(* Logix 5000 project; controller WWTP_CLX vendor 1 type 14 code 54 rev 17.2; software revision 17.00; part 11 of 13 *)

ADD_ON_INSTRUCTION U_FlowTot   (* revision 1.0 *)
// Provides Totalization for Daily & Yearly Flow.
VAR_IN_OUT
   Inp_AIn : P_AIn; {required}   // Flow Analog Input AOI
   Inp_WallClock : U_WallClock; {required}   // PLC Wall Clock
END_VAR
VAR_INPUT
   Inp_ProgStartReq : BOOL := 1;   // Prog Start Request. If needed map to turn on totalizer, (ex. pump running) else Defaults to 1 (always start)
END_VAR
VAR_OUTPUT
   Val_FlowRate : REAL; {visible}   // Current Flow Rate
   Val_DailyTot : REAL; {visible}   // Todays Total Flow
   Val_YestTot : REAL; {visible}   // Yesterday Total Flow
   Val_YearlyTot : REAL; {visible}   // This Year Total Flow
   Val_LastYearTot : REAL; {visible}   // Last Year Total Flow
END_VAR
VAR
   YearlyTotalizer : TOTALIZER := (TimeBase := 3, Gain := 1.0, ProgProgReq := 1, ProgStartReq := 1, OperStartReq := 1, RTSTime := 1, ProgOper := 1, RunStop := 1, TargetFlag := 1, TargetDev1Flag := 1, TargetDev2Flag := 1, DeltaT := 0.010000001);
   DailyTotalizer : TOTALIZER := (TimeBase := 3, Gain := 100000.0, ProgStartReq := 1, OperStartReq := 1, RTSTime := 1, ProgOper := 1, RunStop := 1, TargetFlag := 1, TargetDev1Flag := 1, TargetDev2Flag := 1, DeltaT := 0.010000001);
   FlowRateLowLimit_SSUM : SELECTED_SUMMER := (Gain1 := 1.0, Gain2 := 1.0, Gain3 := 1.0, Gain4 := 1.0, Gain5 := 1.0, Gain6 := 1.0, Gain7 := 1.0, Gain8 := 1.0);
   LowCutoff_BNOT : FBD_BOOLEAN_NOT := (In := 1);
   __l000041A5 : DINT;
   __l000035B4 : REAL;
   __l00000EE7 : BOOL;
   __l00002582 : DINT;
END_VAR

ROUTINE Logic   (* function block diagram *)
   SHEET 1   // Main
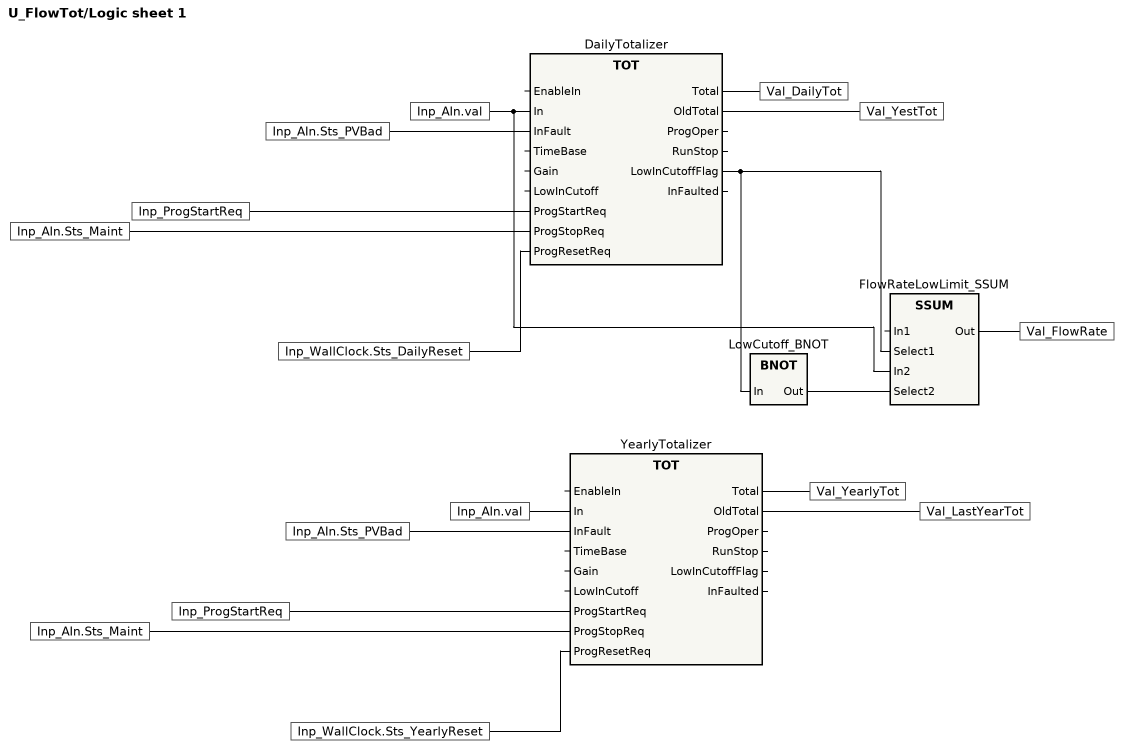
   DailyTotalizer : TOT(In := Inp_AIn.val, InFault := Inp_AIn.Sts_PVBad, ProgStartReq := Inp_ProgStartReq, ProgStopReq := Inp_AIn.Sts_Maint, ProgResetReq := Inp_WallClock.Sts_DailyReset);   // unwired pins: EnableIn TimeBase Gain LowInCutoff ProgOper RunStop InFaulted
   YearlyTotalizer : TOT(In := Inp_AIn.val, InFault := Inp_AIn.Sts_PVBad, ProgStartReq := Inp_ProgStartReq, ProgStopReq := Inp_AIn.Sts_Maint, ProgResetReq := Inp_WallClock.Sts_YearlyReset);   // unwired pins: EnableIn TimeBase Gain LowInCutoff ProgOper RunStop LowInCutoffFlag InFaulted
   LowCutoff_BNOT : BNOT(In := DailyTotalizer.LowInCutoffFlag);
   Val_DailyTot := DailyTotalizer.Total;
   Val_YearlyTot := YearlyTotalizer.Total;
   Val_YestTot := DailyTotalizer.OldTotal;
   FlowRateLowLimit_SSUM : SSUM(Select1 := DailyTotalizer.LowInCutoffFlag, In2 := Inp_AIn.val, Select2 := LowCutoff_BNOT.Out);   // unwired pins: In1
   Val_LastYearTot := YearlyTotalizer.OldTotal;
   Val_FlowRate := FlowRateLowLimit_SSUM.Out;
END_ROUTINE
END_ADD_ON_INSTRUCTION

ADD_ON_INSTRUCTION U_Heartbeat   (* revision 1.0 *)
// Heartbeat Between two PLCs
VAR_INPUT
   CFG_DelayTimerSec : DINT := 30; {visible}   // Delay Timer in Seconds
END_VAR
VAR_OUTPUT
   Heartbeat : BOOL; {visible}   // Heartbeat from Remote PLC
END_VAR
VAR
   DelayTimerOn : TIMER;
   DelayTimerOff : TIMER;
END_VAR

ROUTINE Logic   (* ladder *)
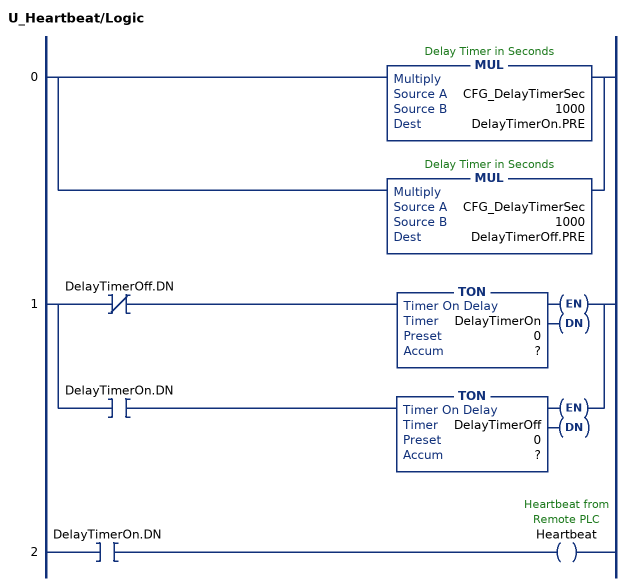
   0: [MUL(CFG_DelayTimerSec,1000,DelayTimerOn.PRE) ,MUL(CFG_DelayTimerSec,1000,DelayTimerOff.PRE) ];
   1: [XIO(DelayTimerOff.DN) TON(DelayTimerOn,?,?) ,XIC(DelayTimerOn.DN) TON(DelayTimerOff,?,?) ];
   2: XIC(DelayTimerOn.DN)OTE(Heartbeat);
END_ROUTINE
END_ADD_ON_INSTRUCTION

ADD_ON_INSTRUCTION U_Module   (* revision 1.0 *)
VAR_INPUT
   EntryStatus : INT; {visible}   // Module Entry Status
   CommLossTimerPresetSec : REAL; {visible}   // Communication Loss Timer Preset (Sec)
END_VAR
VAR_OUTPUT
   CommLoss : BOOL; {visible}   // Communication Loss Alarm
END_VAR
VAR
   ConnectionStatus : DINT;
   CommLossTimer : TIMER := (PRE := 5);
END_VAR

ROUTINE Logic   (* ladder *)
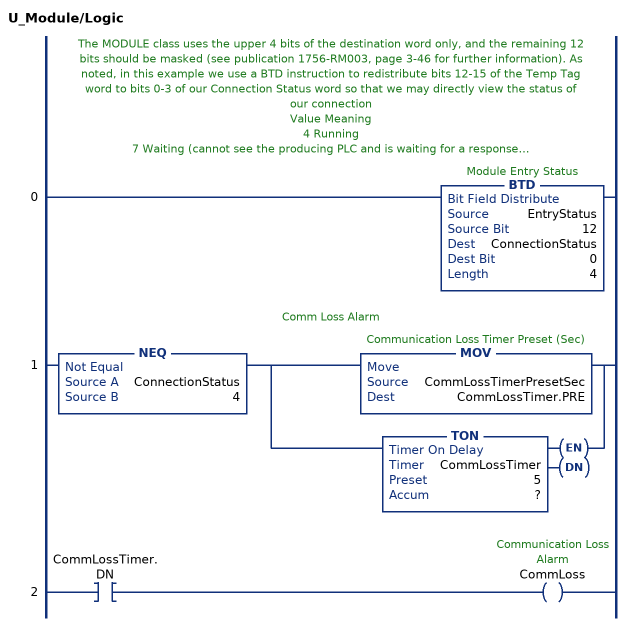
   // The MODULE class uses the upper 4 bits of the destination word only, and the remaining 12 bits should be masked (see publication 1756-RM003, page 3-46 for further information). As noted, in this example we use a BTD instruction to redistribute bits 12-15 of the Temp Tag word to bits 0-3 of our Connection Status word so that we may directly view the status of our connection
   // Value Meaning
   //  4 Running
   //  7 Waiting (cannot see the producing PLC and is waiting for a response)
   //  5 Shutting Down (closing the connection)
   //  1 Faulted (no connection present)
   //  3 Connecting
   // If the connection is good the word will always of value 4. When the connection is lost you will see the value progress to 7, then 5 and finally 1, meaning the connection has faulted and the producing PLC is no longer present.
   0: BTD(EntryStatus,12,ConnectionStatus,0,4);
   // Comm Loss Alarm
   1: NEQ(ConnectionStatus,4)[MOV(CommLossTimerPresetSec,CommLossTimer.PRE) ,TON(CommLossTimer,?,?) ];
   2: XIC(CommLossTimer.DN)OTE(CommLoss);
END_ROUTINE
END_ADD_ON_INSTRUCTION

ADD_ON_INSTRUCTION U_WallClock   (* revision 1.1 *)
// Wall Clock Set time, Current time and Reset bits.
// Revision note:
// Simplified Day of Week calculation, removed unused tags as a result.
VAR_INPUT
   OCmd_SetTime : BOOL; {visible}   // Set the Date and Time Bit
   OSet_Year : DINT; {visible}   // Year To Set
   OSet_Month : DINT; {visible}   // Month To Set
   OSet_Day : DINT; {visible}   // Day To Set
   OSet_Hour : DINT; {visible}   // Hour To Set
   OSet_Minute : DINT; {visible}   // Minute To Set
   OSet_Second : DINT; {visible}   // Second To Set
END_VAR
VAR_OUTPUT
   Val_CurrentYear : DINT; {visible}   // Current Year
   Val_CurrentMonth : DINT; {visible}   // Current Month
   Val_CurrentDay : DINT; {visible}   // Current Day
   Val_CurrentHour : DINT; {visible}   // Current Hour
   Val_CurrentMinute : DINT; {visible}   // Current Minute
   Val_CurrentSecond : DINT; {visible}   // Current Second
   Val_DayOfWeek : DINT; {visible}   // Day of Week 0 = Sun, 1=Mon, 2=Tues, 3=Wed, 4=Thur, 5=Fri, 6=Sat
   Sts_HourlyReset : BOOL; {visible}   // Hourly Reset
   Sts_DailyReset : BOOL; {visible}   // Daily Reset
   Sts_MonthlyReset : BOOL; {visible}   // Monthly Reset
   Sts_YearlyReset : BOOL; {visible}   // Yearly Reset
END_VAR
VAR
   Wrk_SetDateTime : DINT[7];
   Wrk_GetDateTime : DINT[7];   // Result of GSV to Wallclocktime -- input to Day of Week calculation
        [6]   // Microsecond
        [1]   // Month
        [4]   // Minute
        [5]   // Second
        [0]   // Year
        [2]   // Day
        [3]   // Hour
   Wrk_G : DINT;   // Function of Year and Month, used to calculate Day of Week
   Wrk_F : DINT;   // Function of Month, used to calculate Day of Week
   Wrk_DayONS : BOOL;   // One-Shot for daily pulse output
   Wrk_HourONS : BOOL;   // One-Shot for hourly pulse output
   Wrk_MonthONS : BOOL;   // One-Shot for monthly pulse output
   Wrk_YearONS : BOOL;   // One-Shot for yearly pulse output
END_VAR

ROUTINE Logic   (* ladder *)
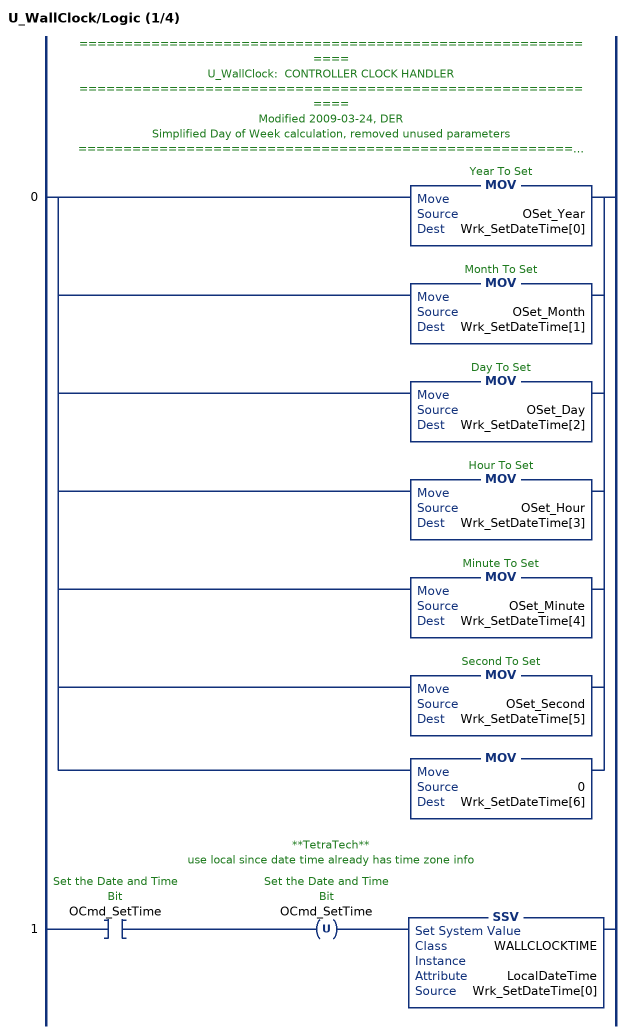
   // ============================================================
   // U_WallClock:  CONTROLLER CLOCK HANDLER
   // ============================================================
   // Modified 2009-03-24, DER
   // Simplified Day of Week calculation, removed unused parameters
   // ============================================================
   // This object manages the controller "Wall Clock", providing date and time services
   // including:
   // * Accepts downloaded date and time and "Set" command from HMI or other sync source and sets the clock
   // * Reads the clock and provides the local date and time to other logic
   // * Calculates and provides the day of the week for the current date
   // * Sets a flag every Hour, Day, Month and Year for resets / data collectors
   // The time is provided as separate Values:
   // Val_CurrentYear : DINT,
   // Val_CurrentMonth : DINT,
   // Val_CurrentDay : DINT,
   // Val_CurrentHour : DINT,
   // Val_CurrentMinute : DINT,
   // Val_CurrentSecond : DINT,
   // Val_DayOfWeek : DINT)
   // ============================================================
   // HANDLE RECEIVED DATE/TIME SYNC, SET CLOCK
   // ============================================================
   // If a date and time have been received with a "Set" command,
   // store the date/time to the controller clock.
   0: [MOV(OSet_Year,Wrk_SetDateTime[0]) ,MOV(OSet_Month,Wrk_SetDateTime[1]) ,MOV(OSet_Day,Wrk_SetDateTime[2]) ,MOV(OSet_Hour,Wrk_SetDateTime[3]) ,MOV(OSet_Minute,Wrk_SetDateTime[4]) ,MOV(OSet_Second,Wrk_SetDateTime[5]) ,MOV(0,Wrk_SetDateTime[6]) ];
   // **TetraTech**
   // use local since date time already has time zone info
   1: XIC(OCmd_SetTime)OTU(OCmd_SetTime)SSV(WALLCLOCKTIME,,LocalDateTime,Wrk_SetDateTime[0]);
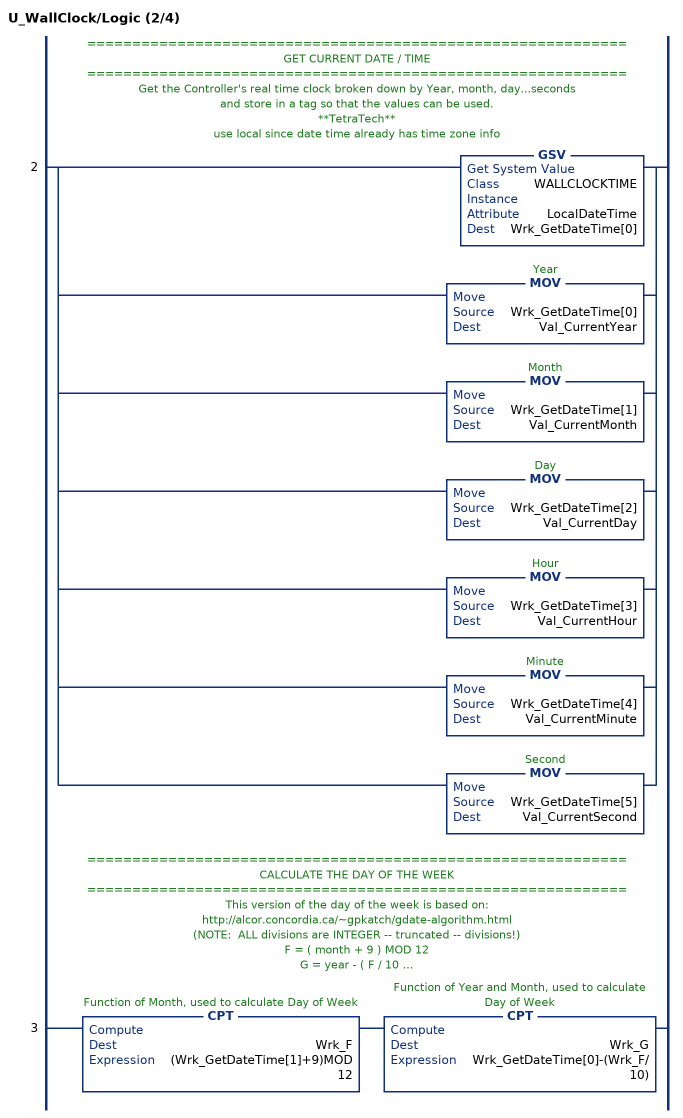
   // ============================================================
   // GET CURRENT DATE / TIME
   // ============================================================
   // Get the Controller's real time clock broken down by Year, month, day...seconds
   // and store in a tag so that the values can be used.
   // **TetraTech**
   // use local since date time already has time zone info
   2: [GSV(WALLCLOCKTIME,,LocalDateTime,Wrk_GetDateTime[0]) ,MOV(Wrk_GetDateTime[0],Val_CurrentYear) ,MOV(Wrk_GetDateTime[1],Val_CurrentMonth) ,MOV(Wrk_GetDateTime[2],Val_CurrentDay) ,MOV(Wrk_GetDateTime[3],Val_CurrentHour) ,MOV(Wrk_GetDateTime[4],Val_CurrentMinute) ,MOV(Wrk_GetDateTime[5],Val_CurrentSecond) ];
   // ============================================================
   // CALCULATE THE DAY OF THE WEEK
   // ============================================================
   // This version of the day of the week is based on:
   // http://alcor.concordia.ca/~gpkatch/gdate-algorithm.html
   // (NOTE:  ALL divisions are INTEGER -- truncated -- divisions!)
   // F = ( month + 9 ) MOD 12
   // G = year - ( F / 10 )
   // Gregorian DayNumber [ D ] = ( 365 * G ) + ( G / 4 ) - ( G / 100 ) + ( G / 400 ) + ( ( ( F * 306 ) + 5 ) / 10 ) + day - 1
   // DayOfWeek = ( DayNumber + 3 ) MOD 7
   // ~~~~~~~~~~~~~~~~~~~~~~~~~~~~~~~~~~~~~~~~~~~~~~~~~~~~~~~~~~~~
   // This rung calculates the "G" and "F" functions shown in the algorithm above.
   // ~~~~~~~~~~~~~~~~~~~~~~~~~~~~~~~~~~~~~~~~~~~~~~~~~~~~~~~~~~~~
   3: CPT(Wrk_F,(Wrk_GetDateTime[1]+9)MOD 12)CPT(Wrk_G,Wrk_GetDateTime[0]-(Wrk_F/10));
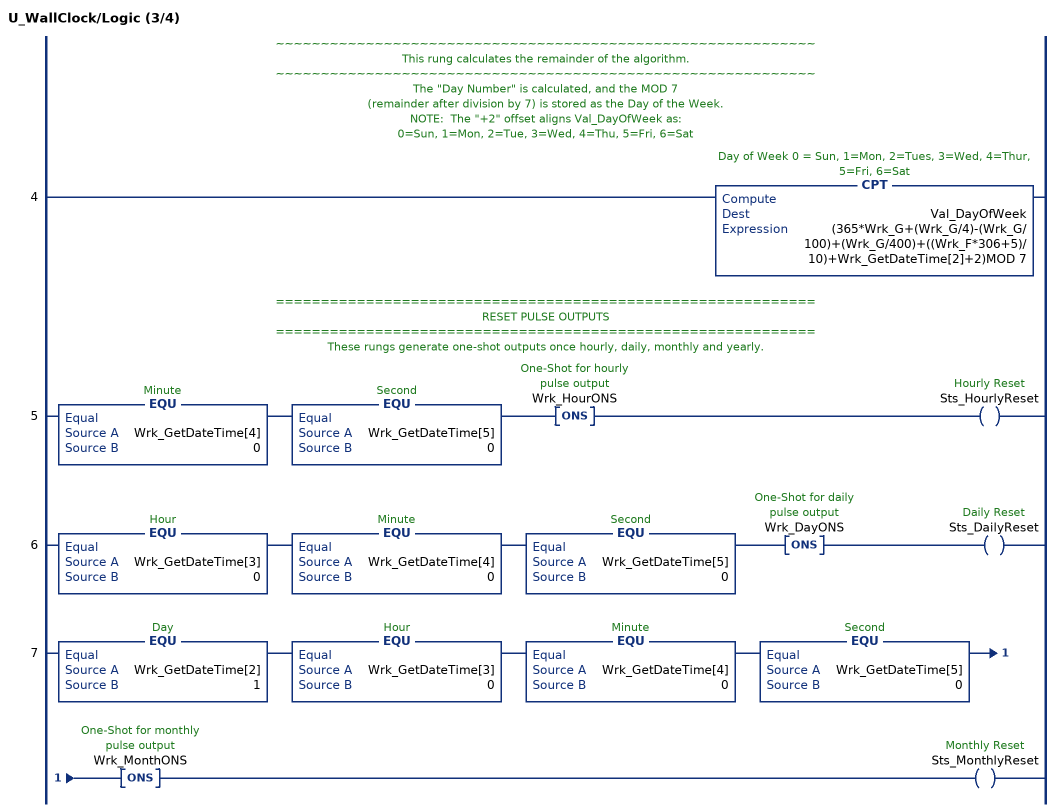
   // ~~~~~~~~~~~~~~~~~~~~~~~~~~~~~~~~~~~~~~~~~~~~~~~~~~~~~~~~~~~~
   // This rung calculates the remainder of the algorithm.
   // ~~~~~~~~~~~~~~~~~~~~~~~~~~~~~~~~~~~~~~~~~~~~~~~~~~~~~~~~~~~~
   // The "Day Number" is calculated, and the MOD 7
   // (remainder after division by 7) is stored as the Day of the Week.
   // NOTE:  The "+2" offset aligns Val_DayOfWeek as:
   // 0=Sun, 1=Mon, 2=Tue, 3=Wed, 4=Thu, 5=Fri, 6=Sat
   4: CPT(Val_DayOfWeek,(365*Wrk_G+(Wrk_G/4)-(Wrk_G/100)+(Wrk_G/400)+((Wrk_F*306+5)/10)+Wrk_GetDateTime[2]+2)MOD 7);
   // ============================================================
   // RESET PULSE OUTPUTS
   // ============================================================
   // These rungs generate one-shot outputs once hourly, daily, monthly and yearly.
   5: EQU(Wrk_GetDateTime[4],0)EQU(Wrk_GetDateTime[5],0)ONS(Wrk_HourONS)OTE(Sts_HourlyReset);
   6: EQU(Wrk_GetDateTime[3],0)EQU(Wrk_GetDateTime[4],0)EQU(Wrk_GetDateTime[5],0)ONS(Wrk_DayONS)OTE(Sts_DailyReset);
   7: EQU(Wrk_GetDateTime[2],1)EQU(Wrk_GetDateTime[3],0)EQU(Wrk_GetDateTime[4],0)EQU(Wrk_GetDateTime[5],0)ONS(Wrk_MonthONS)OTE(Sts_MonthlyReset);
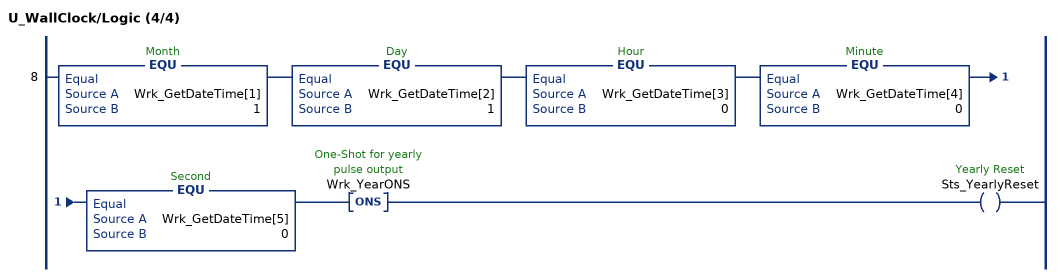
   8: EQU(Wrk_GetDateTime[1],1)EQU(Wrk_GetDateTime[2],1)EQU(Wrk_GetDateTime[3],0)EQU(Wrk_GetDateTime[4],0)EQU(Wrk_GetDateTime[5],0)ONS(Wrk_YearONS)OTE(Sts_YearlyReset);
END_ROUTINE
END_ADD_ON_INSTRUCTION

VAR_GLOBAL   (* controller tags *)
   I_AerTk_InflFlow : REAL := 5.0;
   I_AerTk_InflFlow_IOFault : BOOL;
   I_AlumTk1Lv : ALIAS FOR WWTP_CLX_Rack01_Slot00_CNB:4:I.Ch0Data;
   I_AlumTk1Lv_IOFault : ALIAS FOR WWTP_CLX_Rack01_Slot00_CNB:4:I.Ch0Fault;
   I_FeedP1_Fault : ALIAS FOR WWTP_CLX_Rack01_Slot00_CNB:I.Slot[1].Data.2;
   I_FeedP1_Fault_IOFault : ALIAS FOR WWTP_CLX_Rack01_Slot00_CNB:I.Slot[1].Fault.2;
   I_FeedP1_InAuto : ALIAS FOR WWTP_CLX_Rack01_Slot00_CNB:I.Slot[1].Data.0;
   I_FeedP1_InAuto_IOFault : ALIAS FOR WWTP_CLX_Rack01_Slot00_CNB:I.Slot[1].Fault.0;
   I_FeedP1_OverLoad : ALIAS FOR WWTP_CLX_Rack01_Slot00_CNB:I.Slot[1].Data.3;
   I_FeedP1_OverLoad_IOFault : ALIAS FOR WWTP_CLX_Rack01_Slot00_CNB:I.Slot[1].Fault.3;
   I_FeedP1_RunFdbk : ALIAS FOR WWTP_CLX_Rack01_Slot00_CNB:I.Slot[1].Data.1;
   I_FeedP1_RunFdbk_IOFault : ALIAS FOR WWTP_CLX_Rack01_Slot00_CNB:I.Slot[1].Fault.1;
   I_FeedP1_SpeedFdbk : ALIAS FOR WWTP_CLX_Rack01_Slot00_CNB:4:I.Ch2Data;
   I_FeedP1_SpeedFdbk_IOFault : ALIAS FOR WWTP_CLX_Rack01_Slot00_CNB:4:I.Ch2Fault;
   I_FeedP2_Fault : ALIAS FOR WWTP_CLX_Rack01_Slot00_CNB:I.Slot[1].Data.6;
   I_FeedP2_Fault_IOFault : ALIAS FOR WWTP_CLX_Rack01_Slot00_CNB:I.Slot[1].Fault.6;
   I_FeedP2_InAuto : ALIAS FOR WWTP_CLX_Rack01_Slot00_CNB:I.Slot[1].Data.4;
   I_FeedP2_InAuto_IOFault : ALIAS FOR WWTP_CLX_Rack01_Slot00_CNB:I.Slot[1].Fault.4;
   I_FeedP2_OverLoad : ALIAS FOR WWTP_CLX_Rack01_Slot00_CNB:I.Slot[1].Data.7;
   I_FeedP2_OverLoad_IOFault : ALIAS FOR WWTP_CLX_Rack01_Slot00_CNB:I.Slot[1].Fault.7;
   I_FeedP2_RunFdbk : ALIAS FOR WWTP_CLX_Rack01_Slot00_CNB:I.Slot[1].Data.5;
   I_FeedP2_RunFdbk_IOFault : ALIAS FOR WWTP_CLX_Rack01_Slot00_CNB:I.Slot[1].Fault.5;
   I_FeedP2_SpeedFdbk : ALIAS FOR WWTP_CLX_Rack01_Slot00_CNB:4:I.Ch3Data;
   I_FeedP2_SpeedFdbk_IOFault : ALIAS FOR WWTP_CLX_Rack01_Slot00_CNB:4:I.Ch3Fault;
   LST1_CMPLX_CommFail : U_CommFail := (Inp_Heartbeat := 1, CFG_DelayTimerSec := 60, Sts_CommFail := 1);
   O_FeedP1_Out_Run : ALIAS FOR WWTP_CLX_Rack01_Slot00_CNB:2:O.Data.0;
   O_FeedP1_SpeedRef : ALIAS FOR WWTP_CLX_Rack01_Slot00_CNB:6:O.Ch0Data;
   O_FeedP1_SpeedRef_IOFault : ALIAS FOR WWTP_CLX_Rack01_Slot00_CNB:6:I.Ch0Fault;
   O_FeedP2_Out_Run : ALIAS FOR WWTP_CLX_Rack01_Slot00_CNB:2:O.Data.1;
   O_FeedP2_SpeedRef : ALIAS FOR WWTP_CLX_Rack01_Slot00_CNB:6:O.Ch1Data;
   O_FeedP2_SpeedRef_IOFault : ALIAS FOR WWTP_CLX_Rack01_Slot00_CNB:6:I.Ch1Fault;
   PLC_Device_ResetPB : BOOL;   // Site Wide Device Reset Push Button
   PLC_Heartbeat : U_Heartbeat := (CFG_DelayTimerSec := 1);
   PLC_Simulation : BOOL := 1;   // Application running IN SIMULATION
   PLC_WallClock : U_WallClock := (Val_CurrentYear := 1998, Val_CurrentMonth := 2, Val_CurrentDay := 25, Val_CurrentMinute := 58, Val_CurrentSecond := 30, Val_DayOfWeek := 3);   // Wall Clock
   WWTP_AerTk_InflFlow : UD_Flow := (AIn.Inp_PV := 5.0, AIn.Cfg_SetTrack := 1, AIn.Cfg_PCmdClear := 1, AIn.Cfg_HiHiAckReqd := 1, AIn.Cfg_HiAckReqd := 1, AIn.Cfg_LoAckReqd := 1, AIn.Cfg_LoLoAckReqd := 1, AIn.Cfg_FailAckReqd := 1, AIn.Cfg_HiHiSeverity := 3, AIn.Cfg_HiSeverity := 2, AIn.Cfg_LoSeverity := 2, AIn.Cfg_LoLoSeverity := 3, AIn.Cfg_FailSeverity := 4, AIn.Cfg_InpRawMax := 5.0, AIn.Cfg_PVEUMax := 5.0, AIn.Cfg_HiHiDB := 0.5, AIn.Cfg_HiHiMinDuration := 5, AIn.Cfg_HiDB := 0.5, AIn.Cfg_HiMinDuration := 5, AIn.Cfg_LoDB := 0.5, AIn.Cfg_LoMinDuration := 5, AIn.Cfg_LoLoDB := 0.5, AIn.Cfg_LoLoMinDuration := 5, AIn.Cfg_FailHiLim := 6.0, AIn.Cfg_FailLoLim := -1.0, AIn.Cfg_FailDB := 0.5, AIn.PSet_HiHiLim := 6.0, AIn.PSet_HiLim := 6.0, AIn.PSet_LoLim := -1.0, AIn.PSet_LoLoLim := -1.0, AIn.MSet_SubstPV := 5.0, AIn.OSet_HiHiLim := 6.0, AIn.OSet_HiLim := 6.0, AIn.OSet_LoLim := -1.0, AIn.OSet_LoLoLim := -1.0, AIn.Set_SimPV := 5.0, AIn.Val := 5.0, AIn.Val_InpPV := 5.0, AIn.Val_PVEUMax := 5.0, AIn.Val_HiHiLim := 6.0, AIn.Val_HiLim := 6.0, AIn.Val_LoLim := -1.0, AIn.Val_LoLoLim := -1.0, AIn.Sts_InpPV := 1, AIn.Sts_Oper := 1, AIn.Ack_HiHi := 1, AIn.Ack_Hi := 1, AIn.Ack_Lo := 1, AIn.Ack_LoLo := 1, AIn.Ack_Fail := 1, Tot.Inp_ProgStartReq := 1, Tot.Val_FlowRate := 5.0, Tot.Val_DailyTot := 427429.3, Tot.Val_YestTot := 141377.53, Tot.Val_YearlyTot := 5.9445, Tot.Val_LastYearTot := 8213.769);   // Aeration Tank Influent Flow
   WWTP_Alum : UD_Chemical := (OSet_ChemPercentSolution := 50.0, OSet_ChemWeightLbPGal := 5.0);   // Alum Chemical
   WWTP_AlumTk1Lv : P_AIn := (Inp_PV := 5.0, Inp_PVBad := 1, Cfg_SetTrack := 1, Cfg_PCmdClear := 1, Cfg_HasHiHiAlm := 1, Cfg_HasHiAlm := 1, Cfg_HasLoAlm := 1, Cfg_HasLoLoAlm := 1, Cfg_HiHiAckReqd := 1, Cfg_HiAckReqd := 1, Cfg_LoAckReqd := 1, Cfg_LoLoAckReqd := 1, Cfg_FailAckReqd := 1, Cfg_HiHiSeverity := 3, Cfg_HiSeverity := 2, Cfg_LoSeverity := 2, Cfg_LoLoSeverity := 3, Cfg_FailSeverity := 4, Cfg_InpRawMax := 10.0, Cfg_PVEUMax := 10.0, Cfg_HiHiDB := 1.0, Cfg_HiHiMinDuration := 5, Cfg_HiDB := 1.0, Cfg_HiMinDuration := 5, Cfg_LoDB := 1.0, Cfg_LoMinDuration := 5, Cfg_LoLoDB := 1.0, Cfg_LoLoMinDuration := 5, Cfg_FailHiLim := 1.5e+38, Cfg_FailLoLim := -1.5e+38, PSet_HiHiLim := 9.0, PSet_HiLim := 7.5, PSet_LoLim := 2.5, PSet_LoLoLim := 1.0, MSet_SubstPV := 2.0, OSet_HiHiLim := 9.0, OSet_HiLim := 7.5, OSet_LoLim := 2.5, OSet_LoLoLim := 1.0, Set_SimPV := 5.0, Val := 2.0, Val_InpPV := 5.0, Val_PVEUMax := 10.0, Val_Notify := 4, Val_HiHiLim := 9.0, Val_HiLim := 7.5, Val_LoLim := 2.5, Val_LoLoLim := 1.0, Sts_SubstPV := 1, Sts_Maint := 1, Ack_HiHi := 1, Ack_Hi := 1, Sts_Lo := 1, Alm_Lo := 1, Ack_Lo := 1, Ack_LoLo := 1, Sts_Fail := 1, Ack_Fail := 1, Rdy_InpPV := 1);   // Alum Tank #1 Level
   WWTP_CLX_Rack01_Slot00_Module : U_Module := (EntryStatus := 29184, CommLossTimerPresetSec := 5.0, CommLoss := 1);
   WWTP_FeedP1 : UD_VSD := (Motor.Inp_Ready := 1, Motor.Inp_CommandDir := 1, Motor.Inp_ActualDir := 1, Motor.Inp_FwdPermOK := 1, Motor.Inp_FwdNBPermOK := 1, Motor.Inp_RevPermOK := 1, Motor.Inp_RevNBPermOK := 1, Motor.Inp_IOFault := 1, Motor.Inp_Sim := 1, Motor.Cfg_HasRunFdbk := 1, Motor.Cfg_UseRunFdbk := 1, Motor.Cfg_HasFwdPermObj := 1, Motor.Cfg_HasIntlkObj := 1, Motor.Cfg_HasResInhObj := 1, Motor.Cfg_HasRunTimeObj := 1, Motor.Cfg_SetTrack := 1, Motor.Cfg_HasFailToStartAlm := 1, Motor.Cfg_HasFailToStopAlm := 1, Motor.Cfg_HasIntlkTripAlm := 1, Motor.Cfg_HasDriveFaultAlm := 1, Motor.Cfg_HasIOFaultAlm := 1, Motor.Cfg_FailToStartAckReqd := 1, Motor.Cfg_FailToStopAckReqd := 1, Motor.Cfg_IntlkTripAckReqd := 1, Motor.Cfg_DriveFaultAckReqd := 1, Motor.Cfg_IOFaultAckReqd := 1, Motor.Cfg_FailToStartSeverity := 4, Motor.Cfg_FailToStopSeverity := 4, Motor.Cfg_IntlkTripSeverity := 2, Motor.Cfg_DriveFaultSeverity := 4, Motor.Cfg_IOFaultSeverity := 4, Motor.Cfg_MinSpdRef := 10.0, Motor.Cfg_MaxSpdRef := 100.0, Motor.Cfg_SpeedRefRawMax := 100, Motor.Cfg_SpeedRefEUMax := 100.0, Motor.Cfg_SpeedFdbkRawMax := 100, Motor.Cfg_SpeedFdbkEUMax := 100.0, Motor.Cfg_InpDatalinkRawMax := 4095, Motor.Cfg_InpDatalinkEUMax := 409.5, Motor.Cfg_OutDatalinkMax := 100.0, Motor.Cfg_OutDatalinkRawMax := 4095, Motor.Cfg_OutDatalinkEUMax := 409.5, Motor.Cfg_SimRampT := 10, Motor.Cfg_FailToStartT := 15, Motor.Cfg_FailToStopT := 15, Motor.Cfg_ResetPulseT := 2, Motor.PSet_SpeedRef := 29.803574, Motor.OSet_SpeedRef := 29.803574, Motor.PCmd_Start := 1, Motor.PCmd_Acq := 1, Motor.Val_SpeedRef := 29.803574, Motor.Val_SpeedFdbkEUMax := 100.0, Motor.Val_Notify := 5, Motor.Sts_Stopped := 1, Motor.Sts_CommandDir := 1, Motor.Sts_ActualDir := 1, Motor.Sts_AtSpeed := 1, Motor.Sts_Prog := 1, Motor.Ack_FailToStart := 1, Motor.Ack_FailToStop := 1,
        Motor.Sts_IntlkTrip := 1, Motor.Alm_IntlkTrip := 1, Motor.Ack_DriveFault := 1, Motor.Ack_IOFault := 1, Motor.Rdy_Bypass := 1, Motor.Rdy_Disable := 1, RunTime.Cfg_PCmdClear := 1, RunTime.Val_Starts := 15, RunTime.Val_CurRunHrs := 0.0013933333, RunTime.Val_MaxRunHrs := 17.400898, RunTime.Val_TotRunHrs := 24.5, ResInh.Inp_Stopped := 1, ResInh.Cfg_ThreeColdStarts := 1800, ResInh.Cfg_FirstFailCold := 1800, ResInh.Cfg_SubseqFailCold := 14400, ResInh.Cfg_FirstFailHot := 1800, ResInh.Cfg_SubseqFailHot := 14400, ResInh.Cfg_HotRestartOK := 3600, ResInh.Cfg_RestartHot := 3600, ResInh.Cfg_HotToCold := 57600, ResInh.Val_State := 1, ResInh.Sts_Ready := 1, Intlk.Inp_Intlk00 := 1, Intlk.Cfg_PCmdClear := 1, Intlk.Sts_Intlk := 2#0000_0000_0000_0001, Intlk.Sts_FirstOut := 2#0000_0000_0000_0001, Intlk.Sts_NBFirstOut := 2#0000_0000_0000_0001, Perm.Inp_Perm00 := 1, Perm.Inp_Perm01 := 1, Perm.Inp_Perm02 := 1, Perm.Inp_Perm03 := 1, Perm.Inp_Perm04 := 1, Perm.Inp_Perm05 := 1, Perm.Inp_Perm06 := 1, Perm.Inp_Perm07 := 1, Perm.Inp_Perm08 := 1, Perm.Inp_Perm09 := 1, Perm.Inp_Perm10 := 1, Perm.Inp_Perm11 := 1, Perm.Inp_Perm12 := 1, Perm.Inp_Perm13 := 1, Perm.Inp_Perm14 := 1, Perm.Inp_Perm15 := 1, Perm.Cfg_Bypassable := 2#0000_0000_0000_0001, Perm.Sts_PermOK := 1, Perm.Sts_NBPermOK := 1, Perm.Sts_Perm := 2#1111_1111_1111_1111, Reset.Cfg_MinHoldTime := 1);   // Feed Pump #1
   WWTP_FeedP1_FlowPacing : U_FlowPacing := (Inp_On := 1, OSet_Dosage := 15.0, OSet_PumpCapacityGPH := 35.0, OSet_PumpLength := 100.0, Alm_Prog := 1, Sts_Prog := 1, Rdy_Flow := 1, Sts_PumpStartReqCmd := 1, Val_PumpSpeedRef := 29.803574, Val_PacedFlowMGD := 5.0, Val_ExpectedMaxPacedFlowMGD := 16.776512, Val_ExpectedPumpCapacityGPH := 35.0, Val_ExpectedFlowRateGPH := 10.431251, Val_ChemPercentSolution := 50.0, Val_ChemWeightLbPGal := 5.0);   // Feed Pump #1 Flow Pacing
   WWTP_FeedP1_OverLoad : P_DIn := (Inp_PVBad := 1, Inp_Gate := 1, Cfg_NormTextVis := 1, Cfg_PCmdClear := 1, Cfg_HasTgtDisagreeAlm := 1, Cfg_TgtDisagreeAckReqd := 1, Cfg_TgtDisagreeSeverity := 3, Cfg_TgtDisagreeMinDuration := 5, MSet_SubstPV := 1, Val_Notify := 7, Sts := 1, Sts_SubstPV := 1, Sts_PVBad := 1, Sts_TgtDisagree := 1, Alm_TgtDisagree := 1, Rdy_InpPV := 1);   // Feed Pump #1 Overload
   WWTP_FeedP2 : UD_VSD := (Motor.Inp_Ready := 1, Motor.Inp_CommandDir := 1, Motor.Inp_ActualDir := 1, Motor.Inp_FwdPermOK := 1, Motor.Inp_FwdNBPermOK := 1, Motor.Inp_RevPermOK := 1, Motor.Inp_RevNBPermOK := 1, Motor.Inp_IntlkOK := 1, Motor.Inp_NBIntlkOK := 1, Motor.Inp_IOFault := 1, Motor.Inp_Sim := 1, Motor.Cfg_HasRunFdbk := 1, Motor.Cfg_UseRunFdbk := 1, Motor.Cfg_HasFwdPermObj := 1, Motor.Cfg_HasIntlkObj := 1, Motor.Cfg_HasResInhObj := 1, Motor.Cfg_HasRunTimeObj := 1, Motor.Cfg_SetTrack := 1, Motor.Cfg_HasFailToStartAlm := 1, Motor.Cfg_HasFailToStopAlm := 1, Motor.Cfg_HasIntlkTripAlm := 1, Motor.Cfg_HasDriveFaultAlm := 1, Motor.Cfg_HasIOFaultAlm := 1, Motor.Cfg_FailToStartAckReqd := 1, Motor.Cfg_FailToStopAckReqd := 1, Motor.Cfg_IntlkTripAckReqd := 1, Motor.Cfg_DriveFaultAckReqd := 1, Motor.Cfg_IOFaultAckReqd := 1, Motor.Cfg_FailToStartSeverity := 4, Motor.Cfg_FailToStopSeverity := 4, Motor.Cfg_IntlkTripSeverity := 2, Motor.Cfg_DriveFaultSeverity := 4, Motor.Cfg_IOFaultSeverity := 4, Motor.Cfg_MinSpdRef := 10.0, Motor.Cfg_MaxSpdRef := 100.0, Motor.Cfg_SpeedRefRawMax := 100, Motor.Cfg_SpeedRefEUMax := 100.0, Motor.Cfg_SpeedFdbkRawMax := 100, Motor.Cfg_SpeedFdbkEUMax := 100.0, Motor.Cfg_InpDatalinkRawMax := 4095, Motor.Cfg_InpDatalinkEUMax := 409.5, Motor.Cfg_OutDatalinkMax := 100.0, Motor.Cfg_OutDatalinkRawMax := 4095, Motor.Cfg_OutDatalinkEUMax := 409.5, Motor.Cfg_SimRampT := 10, Motor.Cfg_FailToStartT := 15, Motor.Cfg_FailToStopT := 15, Motor.Cfg_ResetPulseT := 2, Motor.PSet_SpeedRef := 29.383802, Motor.OSet_SpeedRef := 29.383802, Motor.PCmd_Start := 1, Motor.PCmd_Acq := 1, Motor.Val_SpeedRef := 29.383802, Motor.Val_SpeedFdbk := 29.383802, Motor.Val_SpeedFdbkEUMax := 100.0, Motor.Sts_Running := 1, Motor.Sts_CommandDir := 1, Motor.Sts_ActualDir := 1, Motor.Sts_AtSpeed := 1, Motor.Sts_Available := 1,
        Motor.Sts_Prog := 1, Motor.Ack_FailToStart := 1, Motor.Ack_FailToStop := 1, Motor.Ack_IntlkTrip := 1, Motor.Ack_DriveFault := 1, Motor.Ack_IOFault := 1, Motor.Rdy_Bypass := 1, Motor.Rdy_Disable := 1, RunTime.Inp_Running := 1, RunTime.Cfg_PCmdClear := 1, RunTime.Val_Starts := 20, RunTime.Val_CurRunHrs := 0.070049725, RunTime.Val_MaxRunHrs := 0.81247556, RunTime.Val_TotRunHrs := 1.5, ResInh.Inp_Running := 1, ResInh.Cfg_ThreeColdStarts := 1800, ResInh.Cfg_FirstFailCold := 1800, ResInh.Cfg_SubseqFailCold := 30, ResInh.Cfg_FirstFailHot := 1800, ResInh.Cfg_SubseqFailHot := 14400, ResInh.Cfg_HotRestartOK := 3600, ResInh.Cfg_RestartHot := 3600, ResInh.Cfg_HotToCold := 57600, ResInh.Val_State := 3, ResInh.Sts_Ready := 1, Intlk.Cfg_PCmdClear := 1, Intlk.Sts_IntlkOK := 1, Intlk.Sts_NBIntlkOK := 1, Perm.Inp_Perm00 := 1, Perm.Inp_Perm01 := 1, Perm.Inp_Perm02 := 1, Perm.Inp_Perm03 := 1, Perm.Inp_Perm04 := 1, Perm.Inp_Perm05 := 1, Perm.Inp_Perm06 := 1, Perm.Inp_Perm07 := 1, Perm.Inp_Perm08 := 1, Perm.Inp_Perm09 := 1, Perm.Inp_Perm10 := 1, Perm.Inp_Perm11 := 1, Perm.Inp_Perm12 := 1, Perm.Inp_Perm13 := 1, Perm.Inp_Perm14 := 1, Perm.Inp_Perm15 := 1, Perm.Cfg_Bypassable := 2#0000_0000_0000_0001, Perm.Sts_PermOK := 1, Perm.Sts_NBPermOK := 1, Perm.Sts_Perm := 2#1111_1111_1111_1111, Reset.Cfg_MinHoldTime := 1);   // Feed Pump #2
   WWTP_FeedP2_FlowPacing : U_FlowPacing := (Inp_On := 1, OSet_Dosage := 15.0, OSet_PumpCapacityGPH := 35.5, OSet_PumpLength := 100.0, Sts_Prog := 1, Rdy_Flow := 1, Rdy_Pump := 1, Sts_PumpStartReqCmd := 1, Val_PumpSpeedRef := 29.383802, Val_PacedFlowMGD := 5.0, Val_ExpectedMaxPacedFlowMGD := 17.016178, Val_ExpectedPumpCapacityGPH := 35.5, Val_ExpectedFlowRateGPH := 10.43125, Val_ChemPercentSolution := 50.0, Val_ChemWeightLbPGal := 5.0);   // Feed Pump #2 Flow Pacing
   WWTP_FeedP2_OverLoad : P_DIn := (Inp_PVBad := 1, Inp_Gate := 1, Cfg_NormTextVis := 1, Cfg_PCmdClear := 1, Cfg_TgtDisagreeAckReqd := 1, Cfg_TgtDisagreeSeverity := 3, Sts_InpPV := 1, Sts_PVBad := 1, Ack_TgtDisagree := 1, Rdy_SubstPV := 1);   // Feed Pump #2 Overload
   WWTP_FeedSys_OSet_PumpSelect : BOOL := 1;   // Feed Pump System Pump Select
END_VAR

PROGRAM FeedP1   (* main routine Main *)
VAR
   Device : ALIAS FOR WWTP_FeedP1;
   Device_Alm0 : ALIAS FOR WWTP_FeedP1_OverLoad;
   Device_Alm0_Input : ALIAS FOR I_FeedP1_OverLoad;
   Device_Alm0_Input_IOFault : ALIAS FOR I_FeedP1_OverLoad_IOFault;
   Device_Alm1 : P_DIn := (Inp_Gate := 1, Cfg_NormTextVis := 1, Cfg_PCmdClear := 1, Cfg_TgtDisagreeAckReqd := 1, Cfg_TgtDisagreeSeverity := 3, Sts_InpPV := 1, Ack_TgtDisagree := 1, Rdy_SubstPV := 1);
   Device_Alm1_Input : BOOL;
   Device_Alm1_Input_IOFault : BOOL;
   Device_Alm2 : P_DIn := (Inp_Target := 1, Inp_Gate := 1, Cfg_NormTextVis := 1, Cfg_PCmdClear := 1, Cfg_TgtDisagreeAckReqd := 1, Cfg_TgtDisagreeSeverity := 3, Sts_SubstPV := 1, Sts_TgtDisagree := 1, Ack_TgtDisagree := 1, Rdy_InpPV := 1);
   Device_Alm2_Input : BOOL;
   Device_Alm2_Input_IOFault : BOOL;
   Device_Alm3 : P_DIn := (Inp_Target := 1, Inp_Gate := 1, Cfg_NormTextVis := 1, Cfg_PCmdClear := 1, Cfg_TgtDisagreeAckReqd := 1, Cfg_TgtDisagreeSeverity := 3, Sts_SubstPV := 1, Sts_TgtDisagree := 1, Ack_TgtDisagree := 1, Rdy_InpPV := 1);
   Device_Alm3_Input : BOOL;
   Device_Alm3_Input_IOFault : BOOL;
   Device_Alm4 : P_DIn := (Inp_Target := 1, Inp_Gate := 1, Cfg_NormTextVis := 1, Cfg_PCmdClear := 1, Cfg_TgtDisagreeAckReqd := 1, Cfg_TgtDisagreeSeverity := 3, Sts_SubstPV := 1, Sts_TgtDisagree := 1, Ack_TgtDisagree := 1, Rdy_InpPV := 1);
   Device_Alm4_Input : BOOL;
   Device_Alm4_Input_IOFault : BOOL;
   Device_Faulted : ALIAS FOR I_FeedP1_Fault;
   Device_Faulted_IOFault : ALIAS FOR I_FeedP1_Fault_IOFault;
   Device_GroupReset : ALIAS FOR PLC_Device_ResetPB;
   Device_InAuto : ALIAS FOR I_FeedP1_InAuto;
   Device_InAuto_IOFault : ALIAS FOR I_FeedP1_InAuto_IOFault;
   Device_Out_Run : ALIAS FOR O_FeedP1_Out_Run;
   Device_RunFdbk : ALIAS FOR I_FeedP1_RunFdbk;
   Device_RunFdbk_IOFault : ALIAS FOR I_FeedP1_RunFdbk_IOFault;
   Device_SpeedFdbk : ALIAS FOR I_FeedP1_SpeedFdbk;
   Device_SpeedFdbk_IOFault : ALIAS FOR I_FeedP1_SpeedFdbk_IOFault;
   Device_SpeedRef : ALIAS FOR O_FeedP1_SpeedRef;
   Device_SpeedRef_IOFault : ALIAS FOR O_FeedP1_SpeedRef_IOFault;
END_VAR

ROUTINE A01_Alarms   (* ladder *)
// Discrete Alarms
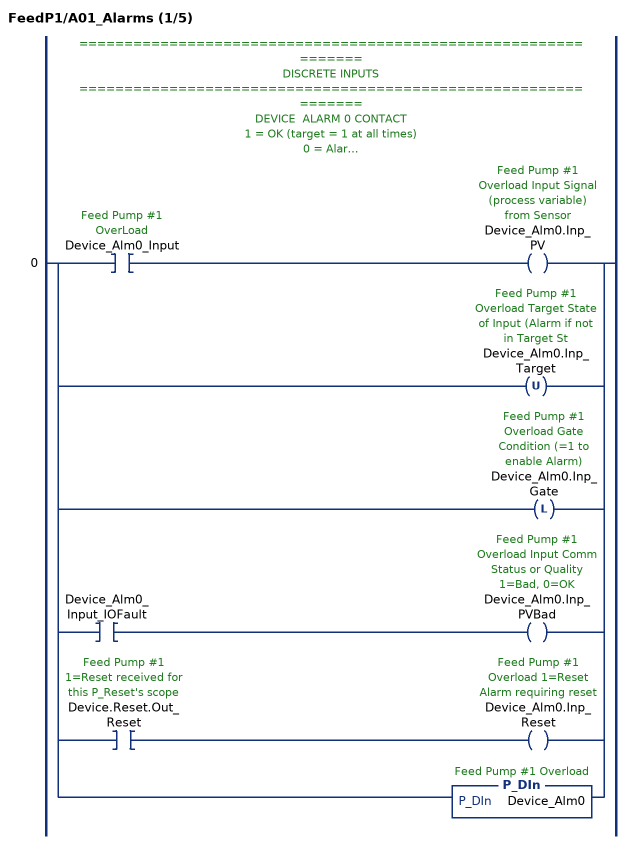
   // ===============================================================
   // DISCRETE INPUTS
   // ===============================================================
   // DEVICE  ALARM 0 CONTACT
   // 1 = OK (target = 1 at all times)
   // 0 = Alarm
   // ALWAYS checked (Gate = 1 at all times)
   0: [XIC(Device_Alm0_Input) OTE(Device_Alm0.Inp_PV) ,OTU(Device_Alm0.Inp_Target) ,OTL(Device_Alm0.Inp_Gate) ,XIC(Device_Alm0_Input_IOFault) OTE(Device_Alm0.Inp_PVBad) ,XIC(Device.Reset.Out_Reset) OTE(Device_Alm0.Inp_Reset) ,P_DIn(Device_Alm0) ];
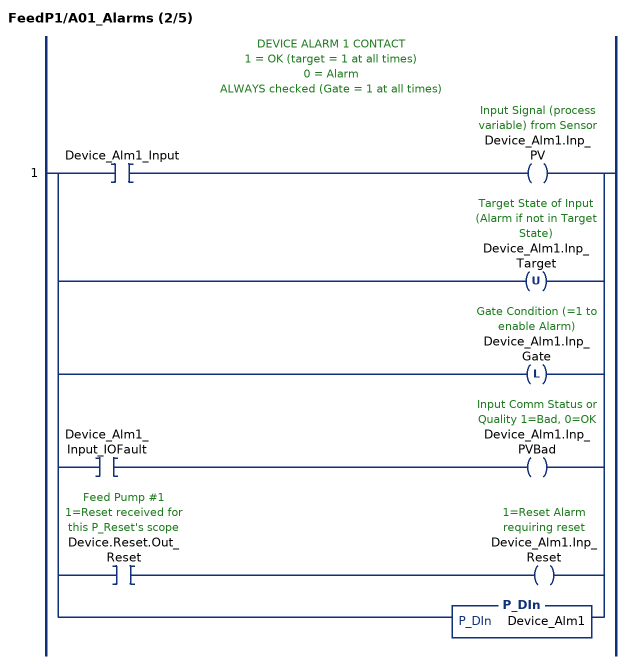
   // DEVICE ALARM 1 CONTACT
   // 1 = OK (target = 1 at all times)
   // 0 = Alarm
   // ALWAYS checked (Gate = 1 at all times)
   1: [XIC(Device_Alm1_Input) OTE(Device_Alm1.Inp_PV) ,OTU(Device_Alm1.Inp_Target) ,OTL(Device_Alm1.Inp_Gate) ,XIC(Device_Alm1_Input_IOFault) OTE(Device_Alm1.Inp_PVBad) ,XIC(Device.Reset.Out_Reset) OTE(Device_Alm1.Inp_Reset) ,P_DIn(Device_Alm1) ];
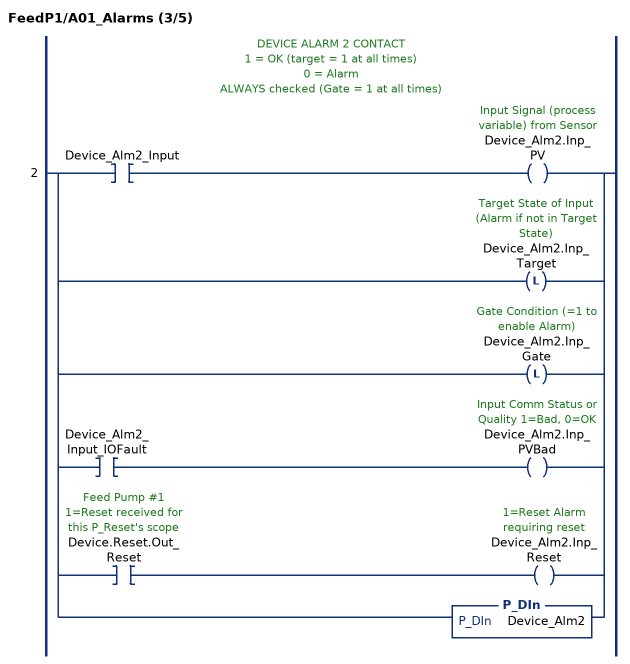
   // DEVICE ALARM 2 CONTACT
   // 1 = OK (target = 1 at all times)
   // 0 = Alarm
   // ALWAYS checked (Gate = 1 at all times)
   2: [XIC(Device_Alm2_Input) OTE(Device_Alm2.Inp_PV) ,OTL(Device_Alm2.Inp_Target) ,OTL(Device_Alm2.Inp_Gate) ,XIC(Device_Alm2_Input_IOFault) OTE(Device_Alm2.Inp_PVBad) ,XIC(Device.Reset.Out_Reset) OTE(Device_Alm2.Inp_Reset) ,P_DIn(Device_Alm2) ];
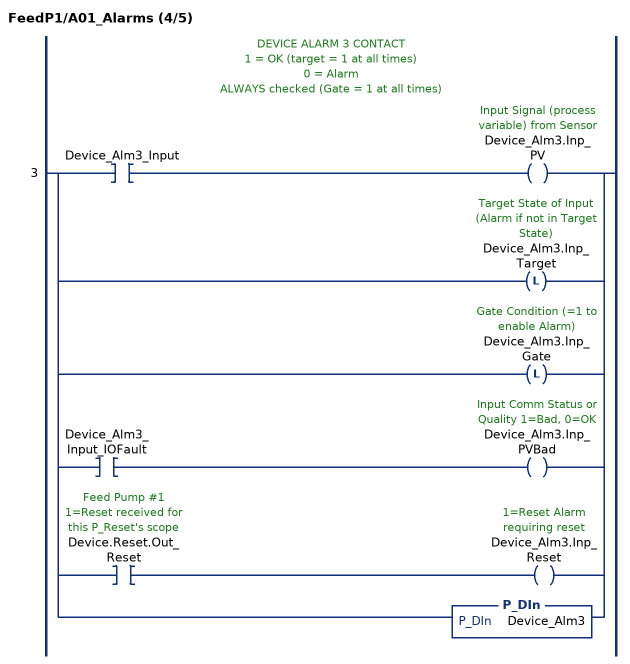
   // DEVICE ALARM 3 CONTACT
   // 1 = OK (target = 1 at all times)
   // 0 = Alarm
   // ALWAYS checked (Gate = 1 at all times)
   3: [XIC(Device_Alm3_Input) OTE(Device_Alm3.Inp_PV) ,OTL(Device_Alm3.Inp_Target) ,OTL(Device_Alm3.Inp_Gate) ,XIC(Device_Alm3_Input_IOFault) OTE(Device_Alm3.Inp_PVBad) ,XIC(Device.Reset.Out_Reset) OTE(Device_Alm3.Inp_Reset) ,P_DIn(Device_Alm3) ];
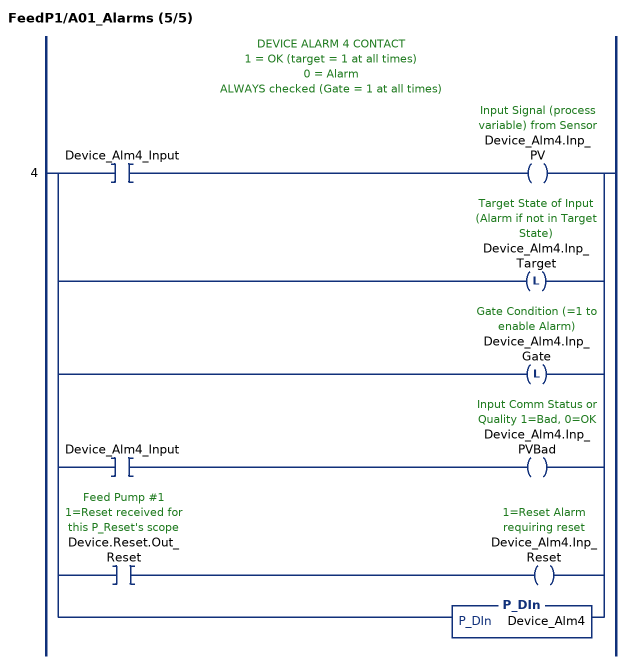
   // DEVICE ALARM 4 CONTACT
   // 1 = OK (target = 1 at all times)
   // 0 = Alarm
   // ALWAYS checked (Gate = 1 at all times)
   4: [XIC(Device_Alm4_Input) OTE(Device_Alm4.Inp_PV) ,OTL(Device_Alm4.Inp_Target) ,OTL(Device_Alm4.Inp_Gate) ,XIC(Device_Alm4_Input) OTE(Device_Alm4.Inp_PVBad) ,XIC(Device.Reset.Out_Reset) OTE(Device_Alm4.Inp_Reset) ,P_DIn(Device_Alm4) ];
END_ROUTINE

ROUTINE A02_Control   (* ladder *)
// Device Contol
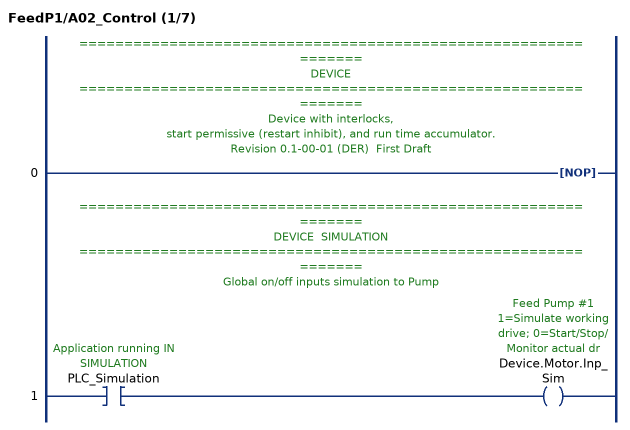
   // ===============================================================
   // DEVICE
   // ===============================================================
   // Device with interlocks,
   // start permissive (restart inhibit), and run time accumulator.
   // Revision 0.1-00-01 (DER)  First Draft
   0: NOP();
   // ===============================================================
   // DEVICE  SIMULATION
   // ===============================================================
   // Global on/off inputs simulation to Pump
   1: XIC(PLC_Simulation)OTE(Device.Motor.Inp_Sim);
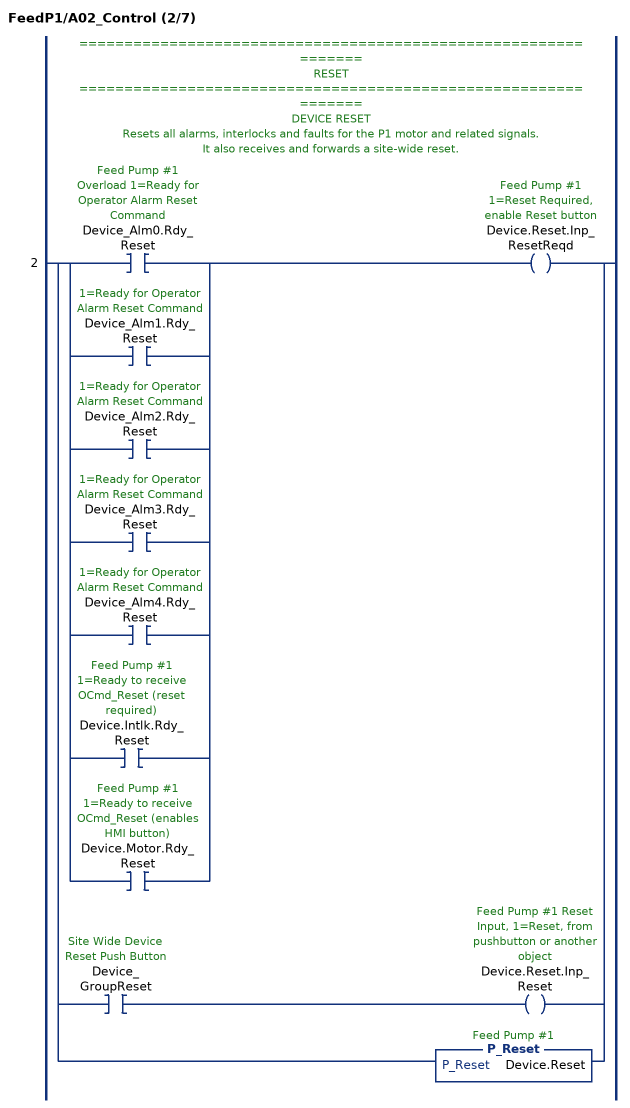
   // ===============================================================
   // RESET
   // ===============================================================
   // DEVICE RESET
   // Resets all alarms, interlocks and faults for the P1 motor and related signals.
   // It also receives and forwards a site-wide reset.
   2: [[XIC(Device_Alm0.Rdy_Reset) ,XIC(Device_Alm1.Rdy_Reset) ,XIC(Device_Alm2.Rdy_Reset) ,XIC(Device_Alm3.Rdy_Reset) ,XIC(Device_Alm4.Rdy_Reset) ,XIC(Device.Intlk.Rdy_Reset) ,XIC(Device.Motor.Rdy_Reset) ] OTE(Device.Reset.Inp_ResetReqd) ,XIC(Device_GroupReset) OTE(Device.Reset.Inp_Reset) ,P_Reset(Device.Reset) ];
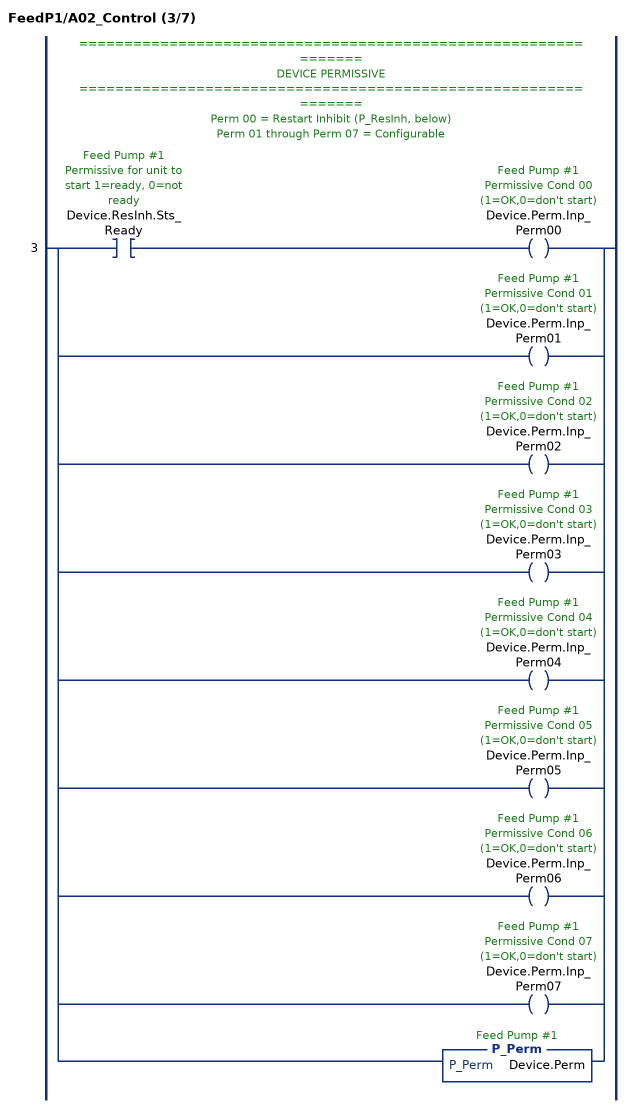
   // ===============================================================
   // DEVICE PERMISSIVE
   // ===============================================================
   // Perm 00 = Restart Inhibit (P_ResInh, below)
   // Perm 01 through Perm 07 = Configurable
   3: [XIC(Device.ResInh.Sts_Ready) OTE(Device.Perm.Inp_Perm00) ,OTE(Device.Perm.Inp_Perm01) ,OTE(Device.Perm.Inp_Perm02) ,OTE(Device.Perm.Inp_Perm03) ,OTE(Device.Perm.Inp_Perm04) ,OTE(Device.Perm.Inp_Perm05) ,OTE(Device.Perm.Inp_Perm06) ,OTE(Device.Perm.Inp_Perm07) ,P_Perm(Device.Perm) ];
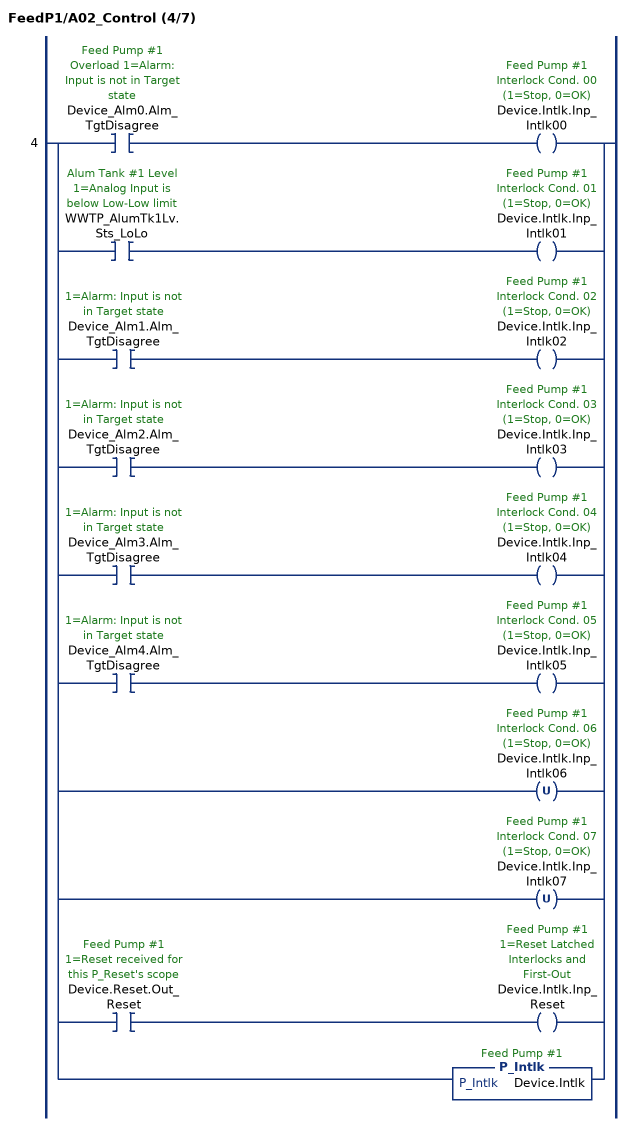
   4: [XIC(Device_Alm0.Alm_TgtDisagree) OTE(Device.Intlk.Inp_Intlk00) ,XIC(WWTP_AlumTk1Lv.Sts_LoLo) OTE(Device.Intlk.Inp_Intlk01) ,XIC(Device_Alm1.Alm_TgtDisagree) OTE(Device.Intlk.Inp_Intlk02) ,XIC(Device_Alm2.Alm_TgtDisagree) OTE(Device.Intlk.Inp_Intlk03) ,XIC(Device_Alm3.Alm_TgtDisagree) OTE(Device.Intlk.Inp_Intlk04) ,XIC(Device_Alm4.Alm_TgtDisagree) OTE(Device.Intlk.Inp_Intlk05) ,OTU(Device.Intlk.Inp_Intlk06) ,OTU(Device.Intlk.Inp_Intlk07) ,XIC(Device.Reset.Out_Reset) OTE(Device.Intlk.Inp_Reset) ,P_Intlk(Device.Intlk) ];
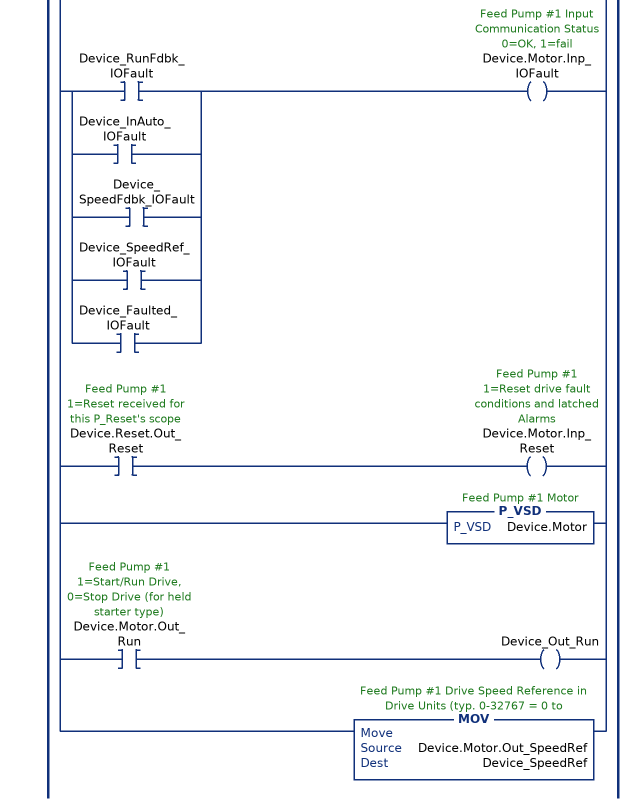
   // ===============================================================
   // DEVICE MOTOR
   // ===============================================================
   // This rung actually monitors and controls the Device motor.
   // Mapping inputs:  Run Feedback
   // Hand Mode selection (local operation)
   // Permissive OK
   // Protective’s OK,
   // I/O Fault signals
   // Pump Reset (above)
   // DEVICE
   // Output Mapping: Starter output
   5: [XIC(Device_RunFdbk) OTE(Device.Motor.Inp_Running) ,MOV(Device_SpeedFdbk,Device.Motor.Inp_SpeedFdbk) ,XIO(Device_InAuto) OTE(Device.Motor.Inp_Hand) ,XIC(Device_Faulted) OTE(Device.Motor.Inp_Faulted) ,XIC(Device.Perm.Sts_PermOK) OTE(Device.Motor.Inp_FwdPermOK) ,XIC(Device.Perm.Sts_NBPermOK) OTE(Device.Motor.Inp_FwdNBPermOK) ,XIC(Device.Intlk.Sts_IntlkOK) OTE(Device.Motor.Inp_IntlkOK) ,XIC(Device.Intlk.Sts_NBIntlkOK) OTE(Device.Motor.Inp_NBIntlkOK) ,[XIC(Device_RunFdbk_IOFault) ,XIC(Device_InAuto_IOFault) ,XIC(Device_SpeedFdbk_IOFault) ,XIC(Device_SpeedRef_IOFault) ,XIC(Device_Faulted_IOFault) ] OTE(Device.Motor.Inp_IOFault) ,XIC(Device.Reset.Out_Reset) OTE(Device.Motor.Inp_Reset) ,P_VSD(Device.Motor) ,XIC(Device.Motor.Out_Run) OTE(Device_Out_Run) ,MOV(Device.Motor.Out_SpeedRef,Device_SpeedRef) ];
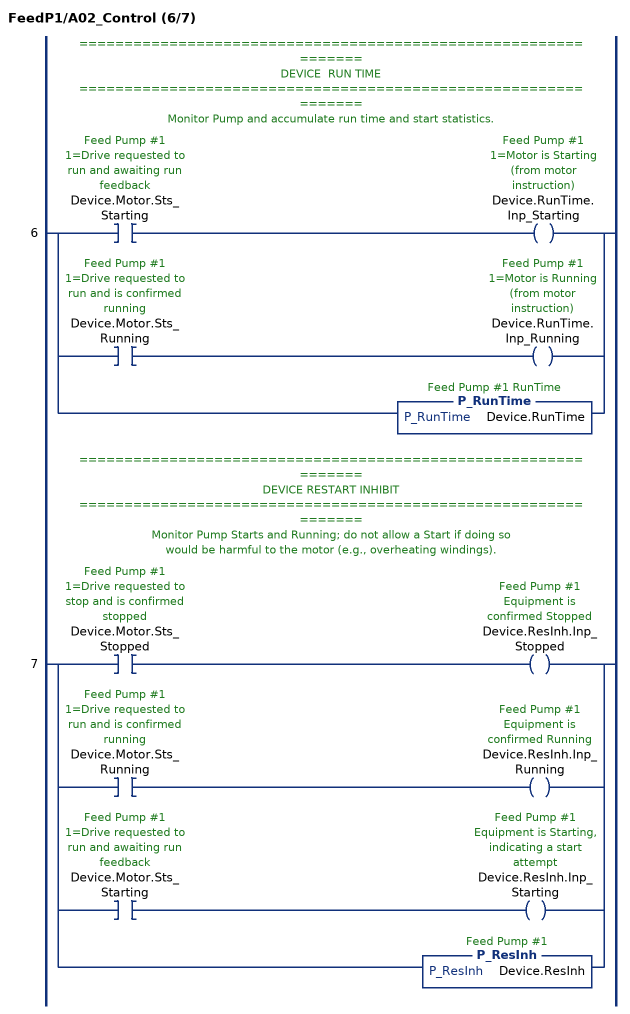
   // ===============================================================
   // DEVICE  RUN TIME
   // ===============================================================
   // Monitor Pump and accumulate run time and start statistics.
   6: [XIC(Device.Motor.Sts_Starting) OTE(Device.RunTime.Inp_Starting) ,XIC(Device.Motor.Sts_Running) OTE(Device.RunTime.Inp_Running) ,P_RunTime(Device.RunTime) ];
   // ===============================================================
   // DEVICE RESTART INHIBIT
   // ===============================================================
   // Monitor Pump Starts and Running; do not allow a Start if doing so
   // would be harmful to the motor (e.g., overheating windings).
   7: [XIC(Device.Motor.Sts_Stopped) OTE(Device.ResInh.Inp_Stopped) ,XIC(Device.Motor.Sts_Running) OTE(Device.ResInh.Inp_Running) ,XIC(Device.Motor.Sts_Starting) OTE(Device.ResInh.Inp_Starting) ,P_ResInh(Device.ResInh) ];
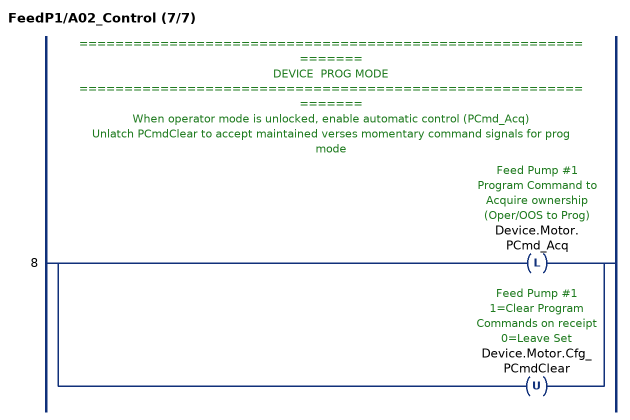
   // ===============================================================
   // DEVICE  PROG MODE
   // ===============================================================
   // When operator mode is unlocked, enable automatic control (PCmd_Acq)
   // Unlatch PCmdClear to accept maintained verses momentary command signals for prog mode
   8: [OTL(Device.Motor.PCmd_Acq) ,OTU(Device.Motor.Cfg_PCmdClear) ];
END_ROUTINE
